DATA_BLOCK "naut_Tags"
{ S7_Optimized_Access := 'TRUE' }
VERSION : 0.1
   VAR
      sel : INT;
      tbl : Array[1..3] of REAL;
   END_VAR

BEGIN
   tbl[1] := 1.0;
   tbl[2] := 2.5;

END_DATA_BLOCK
